SEGMENT_TYPE TestSegment (* Segment with one value *)
  (* Standard: 61499-1; Description: Copyright (c) 2026 Martin Erich Jobst This program and the accompanying materials are made available under the terms of the Eclipse Public License 2.0 which is available at https://www.eclipse.org/legal/epl-2.0/ SPDX-License-Identifier: EPL-2.0 *)
  (* Version 1.0, 2026-10-23, Martin Jobst *)
  {SET_ATTRIBUTE(IntegerAttribute, 15)}
  VAR_INPUT
    VALUE : DINT := DINT#0; (* Segment value *)
  END_VAR
END_SEGMENT_TYPE
